// TIA Portal V15.1 export
// export: Created 2026-11-02T18:55:07.1535265Z, ExportSetting WithDefaults, DisplayName Totally Integrated Automation Portal, DisplayVersion V15.1, DisplayName TIA Portal Openness, DisplayVersion V15.1, DisplayName STEP 7 Professional, DisplayVersion V15.1, DisplayName WinCC Professional, DisplayVersion V15.1
DATA_BLOCK "Sys"   // DB2
{ S7_Optimized_Access := 'TRUE' }
VERSION : 0.1
// stored: AutoNumber false, IsOnlyStoredInLoadMemory false, IsRetainMemResEnabled false, IsWriteProtectedInAS false, MemoryReserve 100
   VAR
      FirstScan : Bool;   // Set by OB100, cleared at the end of Main (C02)
      EStopOK : Bool;   // E-STOP latch: 1 = released and RESET given (C01)
      ResetPulse : Bool;   // RESET S2 rising edge, one scan (R-06)
      ResetMem : Bool;   // RESET edge memory (R-06)
      Alm_EStop : Bool;   // HMI alarm: E-STOP (C01)
      Alm_ParRejected : Bool;   // HMI alarm: a parameter entry was out of range (R-11)
   END_VAR
BEGIN
END_DATA_BLOCK
